(* PLC project Vn_ld_series_parallel, Beckhoff Automation GmbH TwinCAT PLC Control 3.5.13.21 *)
(* stored: creationDateTime 1970-01-01T00:00:00 *)

PROGRAM Vn_ld_series_parallel

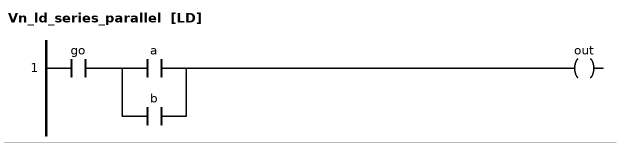
(* LD diagram, written out as Structured Text *)
out := go AND (a OR b);
END_PROGRAM
